FUNCTION_BLOCK "FB_BenchCases"
TITLE = Scenario table and expected values of the test bench (generated)
{ S7_Optimized_Access := 'TRUE' }
AUTHOR : chad416
VERSION : 0.1
//  GENERATED by scripts/make_testbench.py from dmx/bench.py. Do not edit by hand.
//  The expected values are the outcomes of the Python model (dmx/explore.py with the station
//  block in the loop, dmx/ecc200.py for the code content), not of the SCL stand-ins.
//  CaseNo selects the case, PartIx the part inside the case, Row a row of the recipe table.
   VAR_INPUT
      CaseNo : Int;
      PartIx : Int;
      Row : Int;
   END_VAR

   VAR_OUTPUT
      CasesTotal : Int;
      NParts : Int;   // parts in this case
      FaultKind : Int;   // see "FB_SimMarker"; 10 no-read once, 11 no-read always, 12 part taken out, 13 slow record store
      FaultPart : Int;   // the part that gets the fault
      FaultArg : Int;   // fault 12: station step in which the part is taken out
      PartNo : DInt;   // part PartIx of this case
      VarCode : Int;
      RowPartNo : DInt;   // recipe row Row: the job of row n has the number n
      RowVarCode : Int;
      RowJob : Int;
      TmoLoad : Int;   // station time-outs for the bench, in calls
      TmoMark : Int;
      TmoRead : Int;
      TmoRec : Int;
      MaxReads : Int;
      ExpReleased : Int;
      ExpRejected : Int;
      ExpRemoved : Int;
      ExpAlarmSum : Int;
      ExpMarkStarts : Int;
      ExpJobSum : DInt;
      ExpSerialLast : DInt;
      ExpGood : Int;
      ExpVoid : Int;
      ExpRecSerialSum : DInt;
      ExpCodeSum : DInt;
   END_VAR

BEGIN
   #CasesTotal := 21;
   #TmoLoad := 3;
   #TmoMark := 4;
   #TmoRead := 3;
   #TmoRec := 3;
   #MaxReads := 2;

   REGION RecipeRow
   IF #Row >= 1 AND #Row <= 320 THEN
      #RowPartNo := 83700000 + INT_TO_DINT(#Row);
      #RowVarCode := #Row MOD 50;
      #RowJob := #Row;
   ELSE
      #RowPartNo := 0;
      #RowVarCode := 0;
      #RowJob := 0;
   END_IF;
   IF #Row = 205 THEN
      #RowPartNo := 83702051;
      #RowVarCode := 17;
   ELSIF #Row = 206 THEN
      #RowPartNo := 83702052;
      #RowVarCode := 4;
   END_IF;
   END_REGION

   REGION Cases
   #NParts := 0;
   #FaultKind := 0;
   #FaultPart := 0;
   #FaultArg := 0;
   #PartNo := 0;
   #VarCode := 0;
   #ExpReleased := 0;
   #ExpRejected := 0;
   #ExpRemoved := 0;
   #ExpAlarmSum := 0;
   #ExpMarkStarts := 0;
   #ExpJobSum := 0;
   #ExpSerialLast := 0;
   #ExpGood := 0;
   #ExpVoid := 0;
   #ExpRecSerialSum := 0;
   #ExpCodeSum := 0;
   IF #CaseNo = 1 THEN
      // good cycle: parts A
      #NParts := 1;
      #FaultKind := 0;
      #FaultPart := 0;
      #FaultArg := 0;
      IF #PartIx = 1 THEN
         #PartNo := 83702051;
         #VarCode := 17;
      END_IF;
      #ExpReleased := 1;
      #ExpRejected := 0;
      #ExpRemoved := 0;
      #ExpAlarmSum := 0;
      #ExpMarkStarts := 1;
      #ExpJobSum := 205;
      #ExpSerialLast := 1;
      #ExpGood := 1;
      #ExpVoid := 0;
      #ExpRecSerialSum := 1;
      #ExpCodeSum := 10105;
   ELSIF #CaseNo = 2 THEN
      // three part types in a row: parts A B C
      #NParts := 3;
      #FaultKind := 0;
      #FaultPart := 0;
      #FaultArg := 0;
      IF #PartIx = 1 THEN
         #PartNo := 83702051;
         #VarCode := 17;
      ELSIF #PartIx = 2 THEN
         #PartNo := 83702052;
         #VarCode := 4;
      ELSIF #PartIx = 3 THEN
         #PartNo := 83700017;
         #VarCode := 17;
      END_IF;
      #ExpReleased := 3;
      #ExpRejected := 0;
      #ExpRemoved := 0;
      #ExpAlarmSum := 0;
      #ExpMarkStarts := 3;
      #ExpJobSum := 428;
      #ExpSerialLast := 4;
      #ExpGood := 3;
      #ExpVoid := 0;
      #ExpRecSerialSum := 9;
      #ExpCodeSum := 30118;
   ELSIF #CaseNo = 3 THEN
      // changeover back and forth: parts B B A C A
      #NParts := 5;
      #FaultKind := 0;
      #FaultPart := 0;
      #FaultArg := 0;
      IF #PartIx = 1 THEN
         #PartNo := 83702052;
         #VarCode := 4;
      ELSIF #PartIx = 2 THEN
         #PartNo := 83702052;
         #VarCode := 4;
      ELSIF #PartIx = 3 THEN
         #PartNo := 83702051;
         #VarCode := 17;
      ELSIF #PartIx = 4 THEN
         #PartNo := 83700017;
         #VarCode := 17;
      ELSIF #PartIx = 5 THEN
         #PartNo := 83702051;
         #VarCode := 17;
      END_IF;
      #ExpReleased := 5;
      #ExpRejected := 0;
      #ExpRemoved := 0;
      #ExpAlarmSum := 0;
      #ExpMarkStarts := 5;
      #ExpJobSum := 839;
      #ExpSerialLast := 9;
      #ExpGood := 5;
      #ExpVoid := 0;
      #ExpRecSerialSum := 35;
      #ExpCodeSum := 50507;
   ELSIF #CaseNo = 4 THEN
      // part number not in the table, then a good part: parts U A
      #NParts := 2;
      #FaultKind := 0;
      #FaultPart := 0;
      #FaultArg := 0;
      IF #PartIx = 1 THEN
         #PartNo := 12345678;
         #VarCode := 1;
      ELSIF #PartIx = 2 THEN
         #PartNo := 83702051;
         #VarCode := 17;
      END_IF;
      #ExpReleased := 1;
      #ExpRejected := 1;
      #ExpRemoved := 0;
      #ExpAlarmSum := 1;
      #ExpMarkStarts := 1;
      #ExpJobSum := 205;
      #ExpSerialLast := 10;
      #ExpGood := 1;
      #ExpVoid := 0;
      #ExpRecSerialSum := 10;
      #ExpCodeSum := 10104;
   ELSIF #CaseNo = 5 THEN
      // no-read once, second read succeeds: parts A
      #NParts := 1;
      #FaultKind := 10;
      #FaultPart := 1;
      #FaultArg := 0;
      IF #PartIx = 1 THEN
         #PartNo := 83702051;
         #VarCode := 17;
      END_IF;
      #ExpReleased := 1;
      #ExpRejected := 0;
      #ExpRemoved := 0;
      #ExpAlarmSum := 0;
      #ExpMarkStarts := 1;
      #ExpJobSum := 205;
      #ExpSerialLast := 11;
      #ExpGood := 1;
      #ExpVoid := 0;
      #ExpRecSerialSum := 11;
      #ExpCodeSum := 10114;
   ELSIF #CaseNo = 6 THEN
      // no-read on every attempt, then a good part: parts A A
      #NParts := 2;
      #FaultKind := 11;
      #FaultPart := 1;
      #FaultArg := 0;
      IF #PartIx = 1 THEN
         #PartNo := 83702051;
         #VarCode := 17;
      ELSIF #PartIx = 2 THEN
         #PartNo := 83702051;
         #VarCode := 17;
      END_IF;
      #ExpReleased := 1;
      #ExpRejected := 1;
      #ExpRemoved := 0;
      #ExpAlarmSum := 4;
      #ExpMarkStarts := 2;
      #ExpJobSum := 410;
      #ExpSerialLast := 13;
      #ExpGood := 1;
      #ExpVoid := 1;
      #ExpRecSerialSum := 25;
      #ExpCodeSum := 20258;
   ELSIF #CaseNo = 7 THEN
      // marker does not load (time-out), then a good part: parts A A
      #NParts := 2;
      #FaultKind := 1;
      #FaultPart := 1;
      #FaultArg := 0;
      IF #PartIx = 1 THEN
         #PartNo := 83702051;
         #VarCode := 17;
      ELSIF #PartIx = 2 THEN
         #PartNo := 83702051;
         #VarCode := 17;
      END_IF;
      #ExpReleased := 1;
      #ExpRejected := 1;
      #ExpRemoved := 0;
      #ExpAlarmSum := 2;
      #ExpMarkStarts := 1;
      #ExpJobSum := 205;
      #ExpSerialLast := 15;
      #ExpGood := 1;
      #ExpVoid := 1;
      #ExpRecSerialSum := 29;
      #ExpCodeSum := 10154;
   ELSIF #CaseNo = 8 THEN
      // marker hangs without a mark (time-out), then a good part: parts B B
      #NParts := 2;
      #FaultKind := 2;
      #FaultPart := 1;
      #FaultArg := 0;
      IF #PartIx = 1 THEN
         #PartNo := 83702052;
         #VarCode := 4;
      ELSIF #PartIx = 2 THEN
         #PartNo := 83702052;
         #VarCode := 4;
      END_IF;
      #ExpReleased := 1;
      #ExpRejected := 1;
      #ExpRemoved := 0;
      #ExpAlarmSum := 3;
      #ExpMarkStarts := 2;
      #ExpJobSum := 412;
      #ExpSerialLast := 17;
      #ExpGood := 1;
      #ExpVoid := 1;
      #ExpRecSerialSum := 33;
      #ExpCodeSum := 20216;
   ELSIF #CaseNo = 9 THEN
      // marker hangs after a complete mark, then a good part: parts A A
      #NParts := 2;
      #FaultKind := 3;
      #FaultPart := 1;
      #FaultArg := 0;
      IF #PartIx = 1 THEN
         #PartNo := 83702051;
         #VarCode := 17;
      ELSIF #PartIx = 2 THEN
         #PartNo := 83702051;
         #VarCode := 17;
      END_IF;
      #ExpReleased := 1;
      #ExpRejected := 1;
      #ExpRemoved := 0;
      #ExpAlarmSum := 3;
      #ExpMarkStarts := 2;
      #ExpJobSum := 410;
      #ExpSerialLast := 19;
      #ExpGood := 1;
      #ExpVoid := 1;
      #ExpRecSerialSum := 37;
      #ExpCodeSum := 20378;
   ELSIF #CaseNo = 10 THEN
      // marker fault during marking, then a good part: parts A A
      #NParts := 2;
      #FaultKind := 4;
      #FaultPart := 1;
      #FaultArg := 0;
      IF #PartIx = 1 THEN
         #PartNo := 83702051;
         #VarCode := 17;
      ELSIF #PartIx = 2 THEN
         #PartNo := 83702051;
         #VarCode := 17;
      END_IF;
      #ExpReleased := 1;
      #ExpRejected := 1;
      #ExpRemoved := 0;
      #ExpAlarmSum := 3;
      #ExpMarkStarts := 2;
      #ExpJobSum := 410;
      #ExpSerialLast := 21;
      #ExpGood := 1;
      #ExpVoid := 1;
      #ExpRecSerialSum := 41;
      #ExpCodeSum := 20236;
   ELSIF #CaseNo = 11 THEN
      // changeover with a stale job, honest echo: parts A B B
      #NParts := 3;
      #FaultKind := 5;
      #FaultPart := 2;
      #FaultArg := 0;
      IF #PartIx = 1 THEN
         #PartNo := 83702051;
         #VarCode := 17;
      ELSIF #PartIx = 2 THEN
         #PartNo := 83702052;
         #VarCode := 4;
      ELSIF #PartIx = 3 THEN
         #PartNo := 83702052;
         #VarCode := 4;
      END_IF;
      #ExpReleased := 2;
      #ExpRejected := 1;
      #ExpRemoved := 0;
      #ExpAlarmSum := 2;
      #ExpMarkStarts := 2;
      #ExpJobSum := 411;
      #ExpSerialLast := 24;
      #ExpGood := 2;
      #ExpVoid := 1;
      #ExpRecSerialSum := 69;
      #ExpCodeSum := 20225;
   ELSIF #CaseNo = 12 THEN
      // changeover with a stale job, wrong echo: parts A B B
      #NParts := 3;
      #FaultKind := 6;
      #FaultPart := 2;
      #FaultArg := 0;
      IF #PartIx = 1 THEN
         #PartNo := 83702051;
         #VarCode := 17;
      ELSIF #PartIx = 2 THEN
         #PartNo := 83702052;
         #VarCode := 4;
      ELSIF #PartIx = 3 THEN
         #PartNo := 83702052;
         #VarCode := 4;
      END_IF;
      #ExpReleased := 2;
      #ExpRejected := 1;
      #ExpRemoved := 0;
      #ExpAlarmSum := 4;
      #ExpMarkStarts := 3;
      #ExpJobSum := 617;
      #ExpSerialLast := 27;
      #ExpGood := 2;
      #ExpVoid := 1;
      #ExpRecSerialSum := 78;
      #ExpCodeSum := 30397;
   ELSIF #CaseNo = 13 THEN
      // stale serial, honest echo: parts A A A
      #NParts := 3;
      #FaultKind := 7;
      #FaultPart := 2;
      #FaultArg := 0;
      IF #PartIx = 1 THEN
         #PartNo := 83702051;
         #VarCode := 17;
      ELSIF #PartIx = 2 THEN
         #PartNo := 83702051;
         #VarCode := 17;
      ELSIF #PartIx = 3 THEN
         #PartNo := 83702051;
         #VarCode := 17;
      END_IF;
      #ExpReleased := 2;
      #ExpRejected := 1;
      #ExpRemoved := 0;
      #ExpAlarmSum := 2;
      #ExpMarkStarts := 2;
      #ExpJobSum := 410;
      #ExpSerialLast := 30;
      #ExpGood := 2;
      #ExpVoid := 1;
      #ExpRecSerialSum := 87;
      #ExpCodeSum := 20315;
   ELSIF #CaseNo = 14 THEN
      // stale serial, wrong echo: parts A A A
      #NParts := 3;
      #FaultKind := 8;
      #FaultPart := 2;
      #FaultArg := 0;
      IF #PartIx = 1 THEN
         #PartNo := 83702051;
         #VarCode := 17;
      ELSIF #PartIx = 2 THEN
         #PartNo := 83702051;
         #VarCode := 17;
      ELSIF #PartIx = 3 THEN
         #PartNo := 83702051;
         #VarCode := 17;
      END_IF;
      #ExpReleased := 2;
      #ExpRejected := 1;
      #ExpRemoved := 0;
      #ExpAlarmSum := 4;
      #ExpMarkStarts := 3;
      #ExpJobSum := 615;
      #ExpSerialLast := 33;
      #ExpGood := 2;
      #ExpVoid := 1;
      #ExpRecSerialSum := 96;
      #ExpCodeSum := 30426;
   ELSIF #CaseNo = 15 THEN
      // stale job and serial, wrong echo: parts A B A
      #NParts := 3;
      #FaultKind := 9;
      #FaultPart := 2;
      #FaultArg := 0;
      IF #PartIx = 1 THEN
         #PartNo := 83702051;
         #VarCode := 17;
      ELSIF #PartIx = 2 THEN
         #PartNo := 83702052;
         #VarCode := 4;
      ELSIF #PartIx = 3 THEN
         #PartNo := 83702051;
         #VarCode := 17;
      END_IF;
      #ExpReleased := 2;
      #ExpRejected := 1;
      #ExpRemoved := 0;
      #ExpAlarmSum := 4;
      #ExpMarkStarts := 3;
      #ExpJobSum := 616;
      #ExpSerialLast := 36;
      #ExpGood := 2;
      #ExpVoid := 1;
      #ExpRecSerialSum := 105;
      #ExpCodeSum := 30455;
   ELSIF #CaseNo = 16 THEN
      // part taken out during load: parts A A
      #NParts := 2;
      #FaultKind := 12;
      #FaultPart := 1;
      #FaultArg := 30;
      IF #PartIx = 1 THEN
         #PartNo := 83702051;
         #VarCode := 17;
      ELSIF #PartIx = 2 THEN
         #PartNo := 83702051;
         #VarCode := 17;
      END_IF;
      #ExpReleased := 1;
      #ExpRejected := 0;
      #ExpRemoved := 1;
      #ExpAlarmSum := 6;
      #ExpMarkStarts := 1;
      #ExpJobSum := 205;
      #ExpSerialLast := 38;
      #ExpGood := 1;
      #ExpVoid := 1;
      #ExpRecSerialSum := 75;
      #ExpCodeSum := 10202;
   ELSIF #CaseNo = 17 THEN
      // part taken out during marking: parts A A
      #NParts := 2;
      #FaultKind := 12;
      #FaultPart := 1;
      #FaultArg := 40;
      IF #PartIx = 1 THEN
         #PartNo := 83702051;
         #VarCode := 17;
      ELSIF #PartIx = 2 THEN
         #PartNo := 83702051;
         #VarCode := 17;
      END_IF;
      #ExpReleased := 1;
      #ExpRejected := 0;
      #ExpRemoved := 1;
      #ExpAlarmSum := 6;
      #ExpMarkStarts := 2;
      #ExpJobSum := 410;
      #ExpSerialLast := 40;
      #ExpGood := 1;
      #ExpVoid := 1;
      #ExpRecSerialSum := 79;
      #ExpCodeSum := 20343;
   ELSIF #CaseNo = 18 THEN
      // part taken out during read: parts B A
      #NParts := 2;
      #FaultKind := 12;
      #FaultPart := 1;
      #FaultArg := 50;
      IF #PartIx = 1 THEN
         #PartNo := 83702052;
         #VarCode := 4;
      ELSIF #PartIx = 2 THEN
         #PartNo := 83702051;
         #VarCode := 17;
      END_IF;
      #ExpReleased := 1;
      #ExpRejected := 0;
      #ExpRemoved := 1;
      #ExpAlarmSum := 6;
      #ExpMarkStarts := 2;
      #ExpJobSum := 411;
      #ExpSerialLast := 42;
      #ExpGood := 1;
      #ExpVoid := 1;
      #ExpRecSerialSum := 83;
      #ExpCodeSum := 20231;
   ELSIF #CaseNo = 19 THEN
      // part taken out while the record is written: parts A A
      #NParts := 2;
      #FaultKind := 12;
      #FaultPart := 1;
      #FaultArg := 60;
      IF #PartIx = 1 THEN
         #PartNo := 83702051;
         #VarCode := 17;
      ELSIF #PartIx = 2 THEN
         #PartNo := 83702051;
         #VarCode := 17;
      END_IF;
      #ExpReleased := 1;
      #ExpRejected := 0;
      #ExpRemoved := 1;
      #ExpAlarmSum := 6;
      #ExpMarkStarts := 2;
      #ExpJobSum := 410;
      #ExpSerialLast := 44;
      #ExpGood := 2;
      #ExpVoid := 1;
      #ExpRecSerialSum := 130;
      #ExpCodeSum := 20332;
   ELSIF #CaseNo = 20 THEN
      // slow record store: parts A B
      #NParts := 2;
      #FaultKind := 13;
      #FaultPart := 1;
      #FaultArg := 0;
      IF #PartIx = 1 THEN
         #PartNo := 83702051;
         #VarCode := 17;
      ELSIF #PartIx = 2 THEN
         #PartNo := 83702052;
         #VarCode := 4;
      END_IF;
      #ExpReleased := 2;
      #ExpRejected := 0;
      #ExpRemoved := 0;
      #ExpAlarmSum := 0;
      #ExpMarkStarts := 2;
      #ExpJobSum := 411;
      #ExpSerialLast := 46;
      #ExpGood := 2;
      #ExpVoid := 0;
      #ExpRecSerialSum := 91;
      #ExpCodeSum := 20311;
   ELSIF #CaseNo = 21 THEN
      // mixed run of six parts: parts A C B U C A
      #NParts := 6;
      #FaultKind := 0;
      #FaultPart := 0;
      #FaultArg := 0;
      IF #PartIx = 1 THEN
         #PartNo := 83702051;
         #VarCode := 17;
      ELSIF #PartIx = 2 THEN
         #PartNo := 83700017;
         #VarCode := 17;
      ELSIF #PartIx = 3 THEN
         #PartNo := 83702052;
         #VarCode := 4;
      ELSIF #PartIx = 4 THEN
         #PartNo := 12345678;
         #VarCode := 1;
      ELSIF #PartIx = 5 THEN
         #PartNo := 83700017;
         #VarCode := 17;
      ELSIF #PartIx = 6 THEN
         #PartNo := 83702051;
         #VarCode := 17;
      END_IF;
      #ExpReleased := 5;
      #ExpRejected := 1;
      #ExpRemoved := 0;
      #ExpAlarmSum := 1;
      #ExpMarkStarts := 5;
      #ExpJobSum := 650;
      #ExpSerialLast := 51;
      #ExpGood := 5;
      #ExpVoid := 0;
      #ExpRecSerialSum := 245;
      #ExpCodeSum := 50470;
   END_IF;
   END_REGION
END_FUNCTION_BLOCK
